FUNCTION_BLOCK FB_Differential_1
(*
Function block used to calculate differential

Constructor: 		Patryk Panylo
Company:		E. Riexinger GmbH
Date:			05.06.2014
Version:			1.00

Date:			Revision:		Who:				Comment
dd.mm.yyyy		x.xx			Initials			comment

*)
VAR_INPUT
	(* Enummerations *)
	
	(* Variables *)
	bEnable								:BOOL := TRUE;					(* Enable FB *)

	lrInSignal								:LREAL;							(* Input signal *)
	lrDifferentialValue						:LREAL := 1.0;						(* Differential value *)
	lrTaskCycle							:LREAL := 1.0; 					(* Cycle time *)

	(* References *)

	(* Interfaces *)

	(* Instances *)
END_VAR
VAR_OUTPUT
	(* Enummerations *)
	
	(* Variables *)
	lrOutSignal							:LREAL;							(* Output signal *)

	(* References *)

	(* Interfaces *)

	(* Instances *)
END_VAR
VAR
	(* Enummerations *)
	
	(* Variables *)
	bFirstTime							:BOOL;							(* First cycle *)

	lrLastSignal							:LREAL;							(* Last signal *)

	(* References *)

	(* Interfaces *)

	(* Instances *)


END_VAR

IF NOT bEnable
THEN
	lrOutSignal := lrInSignal;

	bFirstTime := FALSE;
	RETURN;
END_IF

IF NOT bFirstTime
THEN
	lrLastSignal := lrInSignal;
	bFirstTime := TRUE;
END_IF

IF lrTaskCycle > 0.0
THEN
	lrOutSignal := lrDifferentialValue * (lrInSignal - lrLastSignal) / lrTaskCycle;
ELSE
	lrOutSignal := 0.0;
END_IF
lrLastSignal := lrInSignal;

END_FUNCTION_BLOCK

(* stored: Version 1.1.0.1, ProductVersion 3.1.4024.15
   POU FB_Differential_1: Id {a478b470-ca5c-41e2-8515-1be507b23dc0}, SpecialFunc None *)
